// TIA Portal V20 export
// export: Created 2026-10-11T05:26:43.4738378Z, ExportSetting WithDefaults, DisplayName Totally Integrated Automation Portal, DisplayVersion V20, DisplayName TIA Portal Openness, DisplayVersion V20, DisplayName TIA Portal Teamcenter Gateway, DisplayVersion V20, DisplayName TIA Portal Version Control Interface, DisplayVersion V20, DisplayName SINAMICS Startdrive Advanced, DisplayVersion V20 SP1 Update 2, DisplayName SINAMICS Startdrive G110M, G120, G120C, G120D, G120P, G115D, DisplayVersion V20 SP1 Update 2, DisplayName SINAMICS Startdrive G130, G150, S120, S150, SINAMICS MV, G220, S200, S210, DisplayVersion V20 SP1 Update 2, DisplayName STEP 7 Professional, DisplayVersion V20, DisplayName STEP 7 Safety, DisplayVersion V20, DisplayName WinCC Basic/Comfort/Advanced, DisplayVersion V20, DisplayName WinCC Professional, DisplayVersion V20, DisplayName WinCC Unified, DisplayVersion V20
FUNCTION "FRK_Start" : Void   // FC14, SCL
{ S7_Optimized_Access := 'TRUE' }
VERSION : 0.1
// stored: AutoNumber true, IsIECCheckEnabled false, SetENOAutomatically false, UDAEnableTagReadback false
   VAR_INPUT
      Supported : Bool;
      Timeout : Time;
      Label : String;
   END_VAR
   VAR_IN_OUT
      Core : "FRK_Core";
      Status : "ST_ModuleStatus";
   END_VAR
BEGIN

   #Core.CommandLabel := #Label;
   IF NOT #Supported THEN
       "FRK_Fault"(Core := #Core,
                   Status := #Status,
                   ReasonCode := 2008,
                   Description := WSTRING#'fraktal.command.unsupported');
   ELSIF #Timeout <= T#0ms THEN
       "FRK_Fault"(Core := #Core,
                   Status := #Status,
                   ReasonCode := 2004,
                   Description := WSTRING#'fraktal.command.timeout.invalid');
   ELSE
       #Core.TimeoutMs := DINT_TO_UDINT(TIME_TO_DINT(#Timeout));
   END_IF;
END_FUNCTION
